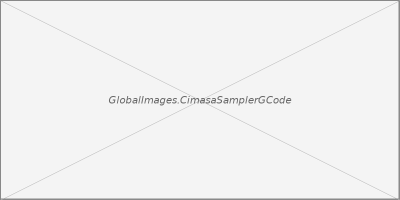
VISUALIZATION V_NCICimasa_SampleBox  // 400x200
    RoundedRectangle (0,0 400x200)
    Image (0,0 400x200), image: GlobalImages.CimasaSamplerGCode
END_VISUALIZATION

(* stored: Version 1.1.0.1, ProductVersion 3.1.4024.15
   Visu V_NCICimasa_SampleBox: Id {4721ca5d-cc2d-45a5-876f-046b5621f450} *)
